Fanuc KAREL source: kb00149.KL

-- PROVISIONAL review KL for V770-1; original PC SHA256 4db1b3d181ccba4b91bd805c62834f05fd01e0dca00e9100ad093daaf786ae5a
-- Incomplete behavior may be omitted. Consult companion uncertainty JSON. Do not deploy.
PROGRAM KB00149
%NOLOCKGROUP
BEGIN
  -- UNRESOLVED_PC offsets 5-12; opcodes 9D,23
  -- UNRESOLVED_PC offsets 17-27; opcodes 27,22,31
  -- UNRESOLVED_PC offsets 32-36; opcodes 7F
END KB00149
